(*
SPDX-FileCopyrightText: © 2026 Oleksandr Tiutyk <trofimich@gmail.com>
SPDX-License-Identifier: MIT
License: https://opensource.org/license/mit
*)

(*!
<summary>Provides fluent assertions on a copied LDATE_AND_TIME value.</summary>
<description>
Copies actual into persistent instance storage before the entry method returns; literals and expression
results therefore remain valid throughout the immediate chain. Owns no heap allocation or pointed-to resource.
The message prefixes every failure until the next preparation. Finish one chain before starting another on
the owning Assertions provider. Use only from the owning test callback on one task, without reentry.
Obtain this context from the owning provider; direct unprepared use is unsupported.
Expected arguments use the declared IEC type; ordinary compiler conversions happen before comparison.
This context does not depend on another assertion context.
Object metadata is available before preparation; inherited equality compares instance identity.
</description>
*)

{attribute 'no_explicit_call' := 'do not call this function block directly'}
FUNCTION_BLOCK LongDateTimeAssertionContext EXTENDS TOF_Core.Object
VAR_STAT
	{attribute 'hide'}
	_ClassName : STRING := __POUNAME();
END_VAR
VAR
	_Actual : LDATE_AND_TIME;
	_TestCase : ITestCase;
	_Message : WSTRING(255);
END_VAR

(*!
<summary>Provides the implementation class name.</summary>
<description>
Borrowed read-only reference to compiler-initialized storage, valid throughout the instance lifetime.
Do not modify the returned reference; no ownership is transferred.
</description>
*)
{attribute 'monitoring' := 'call'}
PROPERTY ClassName : REFERENCE TO STRING
GET
ClassName REF= _ClassName;
END_GET
END_PROPERTY

(*!
<summary>Asserts that the actual value is strictly greater than expected.</summary>
<description>
Records failure without interrupting the callback; preserves the message for the rest of the chain.
</description>
<param name="expected">Expected value converted by the compiler to LDATE_AND_TIME.</param>
*)
METHOD FINAL IsGreaterThan : REFERENCE TO LongDateTimeAssertionContext
VAR_INPUT
	expected : LDATE_AND_TIME;
END_VAR
IF _Actual <= expected THEN
	failComparison(
		expected := expected,
		expectation := "Expected value > "
	);
END_IF

IsGreaterThan REF= THIS^;
END_METHOD

(*!
<summary>Asserts that the actual value meets the inclusive lower boundary.</summary>
<description>
Records failure without interrupting the callback; preserves the message for the rest of the chain.
</description>
<param name="expected">Expected value converted by the compiler to LDATE_AND_TIME.</param>
*)
METHOD FINAL IsGreaterThanOrEquals : REFERENCE TO LongDateTimeAssertionContext
VAR_INPUT
	expected : LDATE_AND_TIME;
END_VAR
IF _Actual < expected THEN
	failComparison(
		expected := expected,
		expectation := "Expected value >= "
	);
END_IF

IsGreaterThanOrEquals REF= THIS^;
END_METHOD

(*!
<summary>Asserts that the actual value is strictly less than expected.</summary>
<description>
Records failure without interrupting the callback; preserves the message for the rest of the chain.
</description>
<param name="expected">Expected value converted by the compiler to LDATE_AND_TIME.</param>
*)
METHOD FINAL IsLessThan : REFERENCE TO LongDateTimeAssertionContext
VAR_INPUT
	expected : LDATE_AND_TIME;
END_VAR
IF _Actual >= expected THEN
	failComparison(
		expected := expected,
		expectation := "Expected value < "
	);
END_IF

IsLessThan REF= THIS^;
END_METHOD

(*!
<summary>Asserts that the actual value meets the inclusive upper boundary.</summary>
<description>
Records failure without interrupting the callback; preserves the message for the rest of the chain.
</description>
<param name="expected">Expected value converted by the compiler to LDATE_AND_TIME.</param>
*)
METHOD FINAL IsLessThanOrEquals : REFERENCE TO LongDateTimeAssertionContext
VAR_INPUT
	expected : LDATE_AND_TIME;
END_VAR
IF _Actual > expected THEN
	failComparison(
		expected := expected,
		expectation := "Expected value <= "
	);
END_IF

IsLessThanOrEquals REF= THIS^;
END_METHOD

(*!
<summary>Provides the library namespace.</summary>
<description>
Borrowed read-only reference to the compiler-initialized namespace, valid throughout the instance lifetime.
Do not modify the returned reference; no ownership is transferred.
</description>
*)
{attribute 'monitoring' := 'call'}
PROPERTY NamespaceName : REFERENCE TO STRING
GET
NamespaceName REF= CurrentNamespace.Name;
END_GET
END_PROPERTY

(*!
<summary>Asserts inequality with the expected value.</summary>
<description>
Records failure without interrupting the callback; preserves the message for the rest of the chain.
</description>
<param name="expected">Expected value converted by the compiler to LDATE_AND_TIME.</param>
*)
METHOD FINAL NotToBe : REFERENCE TO LongDateTimeAssertionContext
VAR_INPUT
	expected : LDATE_AND_TIME;
END_VAR
IF _Actual = expected THEN
	failComparison(
		expected := expected,
		expectation := "Expected value not to be: "
	);
END_IF

NotToBe REF= THIS^;
END_METHOD

(*!
<summary>Copies the actual operand and replaces the chain-wide message.</summary>
<description>
Called by the owning Assertions provider after it verifies the running test case.
No pointer to this method's input storage is retained. The receiver is borrowed until the next preparation;
the owning provider keeps it alive throughout the immediate chain.
</description>
<param name="actual">Value copied into this context.</param>
<param name="testCase">Borrowed failure receiver for the immediate chain.</param>
<param name="message">Copied diagnostic prefix, including empty to clear the previous prefix.</param>
*)
METHOD INTERNAL FINAL Prepare
VAR_INPUT
	actual : LDATE_AND_TIME;
	testCase : ITestCase;
	message : WSTRING(255);
END_VAR
_Actual := actual;
_TestCase := testCase;
_Message := message;
END_METHOD

(*!
<summary>Reports the byte size of this concrete instance.</summary>
<description>
Includes inline fields and nested instances, but excludes separately allocated payloads.
Obtaining the size does not transfer ownership or validate an arbitrary address.
</description>
*)
{attribute 'monitoring' := 'call'}
PROPERTY SelfSize : ULINT
GET
SelfSize := XSIZEOF(THIS^);
END_GET
END_PROPERTY

(*!
<summary>Asserts equality with the expected value.</summary>
<description>
Records failure without interrupting the callback; preserves the message for the rest of the chain.
</description>
<param name="expected">Expected value converted by the compiler to LDATE_AND_TIME.</param>
*)
METHOD FINAL ToBe : REFERENCE TO LongDateTimeAssertionContext
VAR_INPUT
	expected : LDATE_AND_TIME;
END_VAR
IF _Actual <> expected THEN
	failComparison(
		expected := expected,
		expectation := "Expected: "
	);
END_IF

ToBe REF= THIS^;
END_METHOD

(*!
<summary>Formats a failed typed predicate and reports it with the chain message.</summary>
<description>
Does not change operands or chain state. The receiver retains its first failure. Reporting exceptions
propagate to the enclosing test callback handler; an unprepared receiver is a configuration error.
</description>
<param name="expected">Typed expected operand used only for this diagnostic.</param>
<param name="expectation">Prefix identifying the failed predicate.</param>
*)
METHOD PRIVATE failComparison
VAR_INPUT
	expected : LDATE_AND_TIME;
	expectation : WSTRING(40);
END_VAR
VAR
	actualText : WSTRING(255);
	expectedText : WSTRING(255);
	diagnostic : TOF_Core.ERROR_MESSAGE;
END_VAR
actualText := TO_WSTRING(_Actual);
expectedText := TO_WSTRING(expected);

diagnostic := TOF_Core.WideStrings.Concat255(
	expectation,
	expectedText,
	", but was: ",
	actualText
);

TestServices.ReportAssertionFailure(
	testCase := _TestCase,
	message := _Message,
	sourceClassName := ClassName,
	defaultMessage := diagnostic
);
END_METHOD

END_FUNCTION_BLOCK

(* stored: Version 1.1.0.1
   POU LongDateTimeAssertionContext: Id {8cb2268d-8b3b-4529-8e4e-56993ed133d1}, SpecialFunc None
   Folder Service methods: Id {f1e9d44c-a5c7-4e9b-917a-3c46c3b02b45}
   Property ClassName: Id {5bd2e045-3d25-4b46-a6e1-40a4a4a1b8e3}
   Get Get: Id {dc35daa9-f5f2-43d6-bb82-9c9f44a472e3}
   Method IsGreaterThan: Id {07b5a565-3a32-4726-8904-ab0bd9faeaea}
   Method IsGreaterThanOrEquals: Id {af40cccc-0fbf-4384-9eb9-c54aaf1b9201}
   Method IsLessThan: Id {29ba6a00-5e23-4c86-a754-a67ceda5e5d6}
   Method IsLessThanOrEquals: Id {db50ba69-7355-49ad-9ef8-1c5eb8644f68}
   Property NamespaceName: Id {52a7a24b-2000-498d-80de-bdc1664fbcae}
   Get Get: Id {4eca83c7-5904-469d-bffd-5526ba35da35}
   Method NotToBe: Id {e0ef136e-2083-41a8-b865-70900e066766}
   Method Prepare: Id {fa36be80-dc34-45c9-97b4-e5e396b3bc91}
   Property SelfSize: Id {ecc20e91-7492-4ae8-9850-f11b2a4072bc}
   Get Get: Id {8dac0ac5-b8e6-4b40-ae3a-adc0960f7b5a}
   Method ToBe: Id {8e6dfd13-5ad3-4462-89b4-723c00946d7c}
   Method failComparison: Id {6ab38615-d707-4468-8506-469151d0e68f} *)
